Fanuc KAREL source: kb00014.KL

-- PROVISIONAL review KL for V940-1; original PC SHA256 44efd10f0d347bfdd054d5deaf9e4366bf9801e57fd2752fc8311e26bdb8142c
-- Incomplete behavior may be omitted. Consult companion uncertainty JSON. Do not deploy.
PROGRAM KB00014
%NOLOCKGROUP
BEGIN
  -- V9_ZERO_TABLE_METADATA_HINT layout=0002_ascii; no indexed target words; source/name/runtime held
  -- UNRESOLVED_PC offsets 5-21; opcodes 27,22,31,23
  -- UNRESOLVED_PC offsets 26-30; opcodes 7F
END KB00014
